(* IEC 61131-3 sources: modelscript/languages/plcopen/examples/05-automated-bottling-plant, 4 files *)

(* ---- alarm_mgr.st ---- *)
FUNCTION_BLOCK PlantAlarmManager
  VAR_INPUT
    OverPressure : BOOL := FALSE;
    LowTankLevel : BOOL := FALSE;
    AckButton : BOOL := FALSE;
  END_VAR
  VAR_OUTPUT
    AlarmActive : BOOL := FALSE;
    SirenOn : BOOL := FALSE;
  END_VAR

  IF OverPressure OR LowTankLevel THEN
    AlarmActive := TRUE;
    SirenOn := NOT AckButton;
  ELSE
    AlarmActive := FALSE;
    SirenOn := FALSE;
  END_IF;
END_FUNCTION_BLOCK

(* ---- pid_lib.st ---- *)
FUNCTION_BLOCK FillerPressurePid
  VAR_INPUT
    Setpoint : REAL := 2.5;
    ProcessValue : REAL := 2.5;
    Kp : REAL := 1.8;
    Ki : REAL := 0.25;
  END_VAR
  VAR_OUTPUT
    ValveOutputPct : REAL := 0.0;
  END_VAR
  VAR
    Err : REAL := 0.0;
    IntAcc : REAL := 0.0;
  END_VAR

  Err := Setpoint - ProcessValue;
  IntAcc := IntAcc + (Ki * Err * 0.05);
  ValveOutputPct := (Kp * Err) + IntAcc;
  IF ValveOutputPct > 100.0 THEN
    ValveOutputPct := 100.0;
  ELSIF ValveOutputPct < 0.0 THEN
    ValveOutputPct := 0.0;
  END_IF;
END_FUNCTION_BLOCK

(* ---- io_map.st ---- *)
PROGRAM BottlingIoMap
  VAR_INPUT
    RawSensorIn : BOOL := FALSE;
  END_VAR
  VAR_OUTPUT
    MappedBottlePresent : BOOL := FALSE;
  END_VAR

  MappedBottlePresent := RawSensorIn;
END_PROGRAM

(* ---- plant_main.st ---- *)
PROGRAM BottlingPlantMain
  VAR_INPUT
    LineAutoMode : BOOL := TRUE;
    BottleAtFiller : BOOL := FALSE;
    FillerPressureBar : REAL := 2.4;
    EmergencyStop : BOOL := FALSE;
  END_VAR
  VAR_OUTPUT
    MainConveyorRun : BOOL := FALSE;
    FillValveOpen : BOOL := FALSE;
    CapperEngage : BOOL := FALSE;
    BottlesFilled : INT := 0;
  END_VAR
  VAR
    FillDone : BOOL := FALSE;
    FillTimer : TON;
    PressureError : REAL := 0.0;
    TargetPressureBar : REAL := 2.5;
  END_VAR

  IF EmergencyStop THEN
    MainConveyorRun := FALSE;
    FillValveOpen := FALSE;
    CapperEngage := FALSE;
  ELSE
    PressureError := TargetPressureBar - FillerPressureBar;
    MainConveyorRun := LineAutoMode AND NOT BottleAtFiller;
    FillTimer(IN := BottleAtFiller, PT := T#1500ms, Q => FillDone);
    FillValveOpen := BottleAtFiller AND NOT FillDone;
    CapperEngage := FillDone;

    IF FillDone THEN
      BottlesFilled := BottlesFilled + 1;
    END_IF;
  END_IF;
END_PROGRAM
